Fanuc KAREL source: KT00659.KL

PROGRAM KT00659
%NOLOCKGROUP
VAR
  P1: POSITION
  P2: POSITION
  OUT: REAL
BEGIN
  OUT = - P1
END KT00659
